Fanuc KAREL source: kx00011.KL

-- PROVISIONAL review KL for V770-1; original PC SHA256 c5629e7af1593267d29d29cb24ec222e9ac5c6d27ac82684caad8f44cd4df07f
-- Incomplete behavior may be omitted. Consult companion uncertainty JSON. Do not deploy.
PROGRAM KX00011
%NOLOCKGROUP
VAR
  I : INTEGER
  J : INTEGER
  B : BOOLEAN
  F : FILE
  S : STRING[80]
-- UNRESOLVED_DECL P type=000102
BEGIN
  -- UNRESOLVED_PC offsets 5-7; opcodes 9C,65
  -- UNRESOLVED_PC offsets 12-16; opcodes 7F
END KX00011
